(* IEC 61131-3 sources: sis-interlock-demo/src/POUs/Sis/F_VoteCheckCfg, 2 files *)

(* ---- F_VoteCheckCfg.decl.st ---- *)
// Назначение: проверка конфигурации группы голосования: сумма битов VOTE_CFG_* (таблица 4.3);
//             0 — конфигурация верна. Перечисления проверяются сравнениями (строгие перечисления).
// Автор:      kr0nsch
// Версия:     0.1.0
// Документ:   docs/DESIGN.md, раздел «5.9 Проверка конфигурации F_VoteCheckCfg»
// ВНИМАНИЕ:   код демонстрационный и не предназначен для систем безопасности. Реальная ПАЗ
//             требует определения SIL, сертифицированных аппаратных и программных средств
//             и валидации по ГОСТ Р МЭК 61511.
FUNCTION F_VoteCheckCfg : WORD
VAR_IN_OUT CONSTANT
    stCfg : ST_VotingCfg;   // проверяемая конфигурация
END_VAR
VAR
    wErr       : WORD;      // найденные ошибки
    uiN        : UINT;      // каналов в схеме; 0 — схема неверна
    xBypassBad : BOOL;      // недопустимое число байпасов
END_VAR

(* ---- F_VoteCheckCfg.impl.st ---- *)
wErr := 0;
uiN := F_VoteArchChannels(eArch := stCfg.eArch);

// Схема: только 1oo1, 1oo2, 2oo2, 2oo3 (None и ForcedTrip — ошибка)
IF uiN = 0 THEN
    wErr := wErr OR GVL_Const.VOTE_CFG_ARCH;
END_IF

IF NOT (stCfg.ePolicy = E_DegradePolicy.VoteTrip OR stCfg.ePolicy = E_DegradePolicy.DegradeSafe
    OR stCfg.ePolicy = E_DegradePolicy.DegradeAvailable)
THEN
    wErr := wErr OR GVL_Const.VOTE_CFG_POLICY;
END_IF

IF NOT (stCfg.eInput = E_SisInputKind.Discrete OR stCfg.eInput = E_SisInputKind.Analog) THEN
    wErr := wErr OR GVL_Const.VOTE_CFG_INPUT;
END_IF

// Поля аналога проверяются только для Analog; для Discrete они не действуют
IF stCfg.eInput = E_SisInputKind.Analog THEN
    IF NOT PL.F_IsFinite(rIn := stCfg.rTripLimit_eu) OR NOT PL.F_IsFinite(rIn := stCfg.rHyst_eu)
        OR stCfg.rHyst_eu < 0.0
        OR NOT (stCfg.eLimitDir = E_LimitDir.High OR stCfg.eLimitDir = E_LimitDir.Low)
    THEN
        wErr := wErr OR GVL_Const.VOTE_CFG_LIMIT;
    END_IF
    IF NOT PL.F_IsFinite(rIn := stCfg.rDiscrepancyMax_eu) OR stCfg.rDiscrepancyMax_eu < 0.0
        OR stCfg.tDiscrepancyDelay > GVL_Const.SIS_DELAY_MAX
    THEN
        wErr := wErr OR GVL_Const.VOTE_CFG_DISCREPANCY;
    END_IF
END_IF

// Байпасов — не больше N − 1 (хотя бы один канал голосует); при неверной схеме — ни одного
IF uiN = 0 THEN
    xBypassBad := stCfg.uiMaxBypass > 0;
ELSE
    xBypassBad := stCfg.uiMaxBypass > uiN - 1;
END_IF
IF xBypassBad OR stCfg.tBypassMax > GVL_Const.SIS_BYPASS_MAX THEN
    wErr := wErr OR GVL_Const.VOTE_CFG_BYPASS;
END_IF

F_VoteCheckCfg := wErr;
